FUNCTION_BLOCK F (* Positive: an input override reaches one state from every position, and not all scans pass through it *)
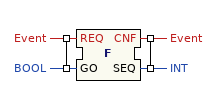
  EVENT_INPUT
    REQ WITH GO;
  END_EVENT
  EVENT_OUTPUT
    CNF WITH SEQ;
  END_EVENT
  VAR_INPUT
    GO : BOOL;
  END_VAR
  VAR_OUTPUT
    SEQ : INT;
  END_VAR
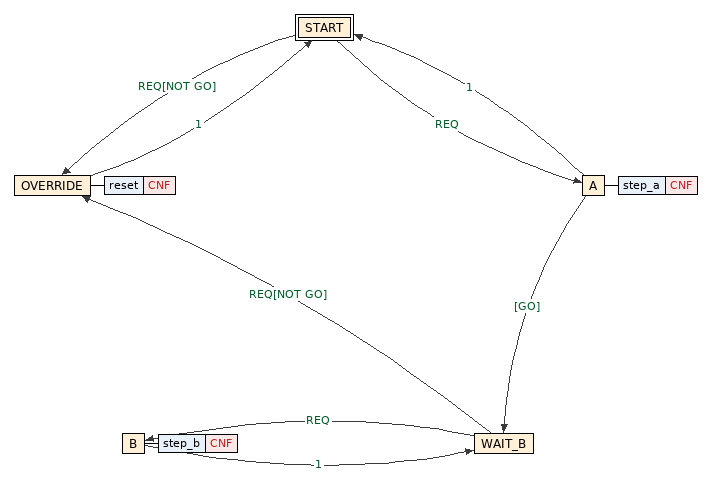
  EC_STATES
    START;
    A : step_a -> CNF;
    WAIT_B;
    B : step_b -> CNF;
    OVERRIDE : reset -> CNF;
  END_STATES
  EC_TRANSITIONS
    START TO OVERRIDE := REQ[NOT GO];
    START TO A := REQ;
    A TO WAIT_B := [GO];
    A TO START := 1;
    WAIT_B TO OVERRIDE := REQ[NOT GO];
    WAIT_B TO B := REQ;
    B TO WAIT_B := 1;
    OVERRIDE TO START := 1;
  END_TRANSITIONS
  ALGORITHM step_a IN ST:
SEQ := 0;
IF GO THEN
  SEQ := 1;
END_IF;
  END_ALGORITHM
  ALGORITHM step_b IN ST:
IF NOT GO THEN
  SEQ := 0;
END_IF;
  END_ALGORITHM
  ALGORITHM reset IN ST:
SEQ := 0;
  END_ALGORITHM
END_FUNCTION_BLOCK
